Fanuc KAREL source: kd00025.KL

-- PROVISIONAL review KL for V940-1; original PC SHA256 f76e3cb649905f0adcbbf208b76ed8566756cdda2c5491325f7354b2c626c7f1
-- Incomplete behavior may be omitted. Consult companion uncertainty JSON. Do not deploy.
PROGRAM KD00025
%NOLOCKGROUP
VAR
  I : INTEGER
  J : INTEGER
  B : BOOLEAN
  R : REAL
  S : STRING[80]
BEGIN
  -- V9_ZERO_TABLE_METADATA_HINT layout=0001; no indexed target words; source/name/runtime held
  -- UNRESOLVED_PC offsets 5-31; opcodes 9D,2E,25,81,18,9D,1B,9D,12,22,9D,13,04
  -- UNRESOLVED_PC offsets 36-40; opcodes 7F
END KD00025
